FUNCTION_BLOCK Button_IMC (* Extracted Composite Function Block Type *)
  (* Standard: 61499-2 *)
  (* Version 10/27/2026, lizar *)
  PACKAGE Main;
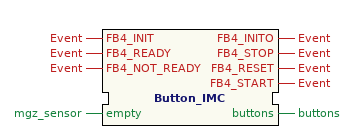
  EVENT_INPUT
    FB4_INIT; (* Event input *)
    FB4_READY;
    FB4_NOT_READY;
  END_EVENT
  EVENT_OUTPUT
    FB4_INITO;
    FB4_STOP;
    FB4_RESET;
    FB4_START;
  END_EVENT
  SOCKETS
    empty : mgz_sensor;
  END_SOCKETS
  PLUGS
    buttons : buttons;
  END_PLUGS
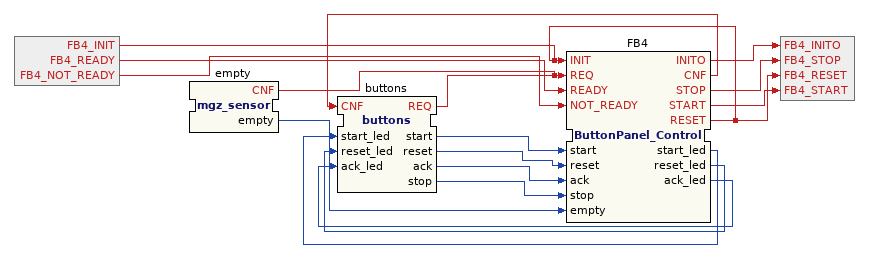
  FBS
    FB4 : ButtonPanel_Control;
  END_FBS
  EVENT_CONNECTIONS
    FB4.RESET TO FB4.INIT;
    FB4_INIT TO FB4.INIT;
    FB4_READY TO FB4.READY;
    FB4_NOT_READY TO FB4.NOT_READY;
    FB4.INITO TO FB4_INITO;
    FB4.STOP TO FB4_STOP;
    FB4.RESET TO FB4_RESET;
    FB4.START TO FB4_START;
    buttons.REQ TO FB4.REQ;
    FB4.CNF TO buttons.CNF;
    empty.CNF TO FB4.REQ;
  END_CONNECTIONS
  DATA_CONNECTIONS
    buttons.start TO FB4.start;
    buttons.reset TO FB4.reset;
    buttons.ack TO FB4.ack;
    buttons.stop TO FB4.stop;
    FB4.start_led TO buttons.start_led;
    FB4.reset_led TO buttons.reset_led;
    FB4.ack_led TO buttons.ack_led;
    empty.empty TO FB4.empty;
  END_CONNECTIONS
END_FUNCTION_BLOCK
